// SIMATIC S7-200 project (STEP 7-Micro/WIN), CPU 226 CN REL 02.01

SYMBOL_TABLE ????1
SI1              I0.0     // Sensor de riel
FCI              I0.1     // Final de carrera derecha
FCF              I0.2     // Final de carrera izquierda
SM2B             I0.4     // Sensor de elevamiento vertical
SM2A             I0.3     // Sensor retraido vertical
SAH              I0.5     // Sensor antiHorario de giro
SH               I0.6     // Sensor Horario de giro
SM3B             I0.7     // Sesor extendido horizontal
SM3A             I1.0     // Sensor retraido horizontal
SM4C             I1.1     // Sensor Garra cerrada
                 I1.3     // Alarma servo
SB_2             I2.4     // Pulsador de parada
SB_1             I2.5     // Pulsador de marcha
QS               I2.6     // Zeta de emergencia
SA               I2.7     // Selector de modo
PULSO            Q0.0     // Pulso
DIR              Q0.1     // Direccion
KV2              Q0.3     // Cilndro neumatico vertical
KV1A             Q0.4     // Cilindro rotarorio anti horario
KV1H             Q0.5     // Cilindro rotatorio horario
KV3              Q0.6     // Cilindro doble horizontal
KV4C             Q0.7     // Garra cerrada
KV4A             Q1.0     // Garra abierta
HL1              Q1.5     // Piloto Amarillo
HL2              Q1.6     // Piloto Verde
HL3              Q1.7     // Piloto Rojo
E0               M0.0     // Estado 0
E1               M0.1     // Estado 1
E2               M0.2
E3               M0.3
E4               M0.4
E5               M0.5
E6               M0.6
E7               M0.7
E8               M1.0
E9               M1.1
E10              M1.2
E11              M1.3
E12              M1.4
E13              M1.5
E14              M1.6
E15              M1.7
E16              M2.0
E17              M2.1
E18              M2.2
E19              M2.3
E20              M2.4
E21              M2.5
E22              M2.6
E23              M2.7
EP               M3.0     // Estado de parada momentanea
Marca            M3.1     // Marca auxiliar
EM               M3.2     // Estado de emergencia
SB1_UT           M4.0     // Pulsador de marcha
SB2_UT           M4.1     // Pulsador de parada
QS_UT            M4.2     // Zeta de emergencia
POS_UA           M5.0     // Posicionamiento a la Unidad de Alimentacion
POS_UE           M5.1     // Posicionamiento a la Unidad de Ensamblaje
POS_UP           M5.2     // Posicionamiento a la Unidad de Procesamiento
POS_US           M5.3     // Posicionamiento a la Unidad de Seleccion
END_UA           V0.0     // Finializacion de la Unidad de Alimentacion
END_UE           V12.0    // Finalizacion de la Unidad de Ensamblaje
END_UP           V6.0     // Finalizacion de la Unidad de Procesamiento
END_US           V18.0    // Finalizacion de la Unidad de Seleccion
IN_UA            V3.0     // Iniciar Unidad de Alimentacion
IN_UE            V15.0    // Iniciar Unidad de Ensamblaje
IN_UP            V9.0     // Iniciar Unidad de Procesamiento
IN_US            V21.0    // Iniciar Unidad de Seleccion
                          // UNIDAD DE ALIMENTACION
SB1_UA           M4.3     // Pulsador de marcha
SB2_UA           M4.4     // Pulsador de parada
QS_UA            M4.5     // Zeta de emergencia
KV1_UA           V0.1     // Cilindro neumatico Retenedor
KV2_UA           V0.2     // Cilindro neumatico de empuje
SF_UA            V0.3     // Sensor Fotoelectrico Final
SP_UA            V0.4     // Sensor Fotoelectrico Superior
SP1_UA           V0.5     // Sensor Fotoelectrico Inferior
HL1_UA           V0.6     // Piloto de parada
HL2_UA           V0.7     // Piloto de marcha
HL3_UA           V1.0     // Piloto de emergencia
                          // UNIDAD DE ENSAMBLAJE
SB1_UE           M15.1    // Pulsador de marcha
SB2_UE           M15.2    // Pulsador de parada
QS_UE            M15.3    // Zeta de emergencia
KV1_UE           V12.1    // Cilindro liberador
KV2_UE           V12.2    // Cildro sujetador
KV3_UE           V12.3    // Cilindro rotatorio
KV4_UE           V12.4    // Cilindro vertical
KV5_UE           V12.5    // Cilindro horizontal
KV6_UE           V12.6    // Cilindro de garra
SP1_UE           V13.0    // Sensor del tubo inferior
SP_UE            V13.1    // Sensor del tubo superiro
SST_UE           V13.2    // Sensor salida del tubo
SG_UE            V13.3    // Sensor de recogida de pieza
SF_UE            V13.4    // Sensor de posicion de pieza grande
HL1_UE           V13.5    // Piloto de parada
HL2_UE           V13.6    // Piloto de marcha
HL3_UE           V13.7    // Piloto de emergencia
                          // UNIDAD DE PROCESAMIENTO
SB1_UP           M9.1     // Pulsador de marcha
SB2_UP           M9.2     // Pulsador de parada
QS_UP            M9.3     // Zeta de emergencia
KV1_UP           V6.1     // Cilindro neumatico horizontal
KV2_UP           V6.2     // Cilindro de la pinza
KV3_UP           V6.3     // Cilindro neumatico de compresion
SF1_UP           V6.4     // Sensor optico
HL1_UP           V6.5     // Piloto de parada
HL2_UP           V6.6     // Piloto de marcha
HL3_UP           V6.7     // Piloto de emergencia
                          // UNIDAD DE SELECCION
SB1_US           M21.1    // Pulsador de marcha
SB2_US           M21.2    // Pulsador de parada
QS_US            M21.3    // Zeta de emergencia
KV1_US           V18.1    // Cilindro neumatico 1
KV2_US           V18.2    // Cilindro neumatico 2
KV3_US           V18.3    // Cilindro neumatico 3
motor            V18.4    // Motor
SF_US            V18.5    // Sensor de objetos
SII_US           V18.6    // Sensor inductivo (Metal)
SP_US            V18.7    // Sensor magnetico (plastico)
HL1_US           V19.0    // Piloto de parada
HL2_US           V19.1    // Piloto de marcha
HL3_US           V19.2    // Piloto de emergencia
END_SYMBOL_TABLE

ORGANIZATION_BLOCK PRINCIPAL:OB1
TITLE=????
BEGIN
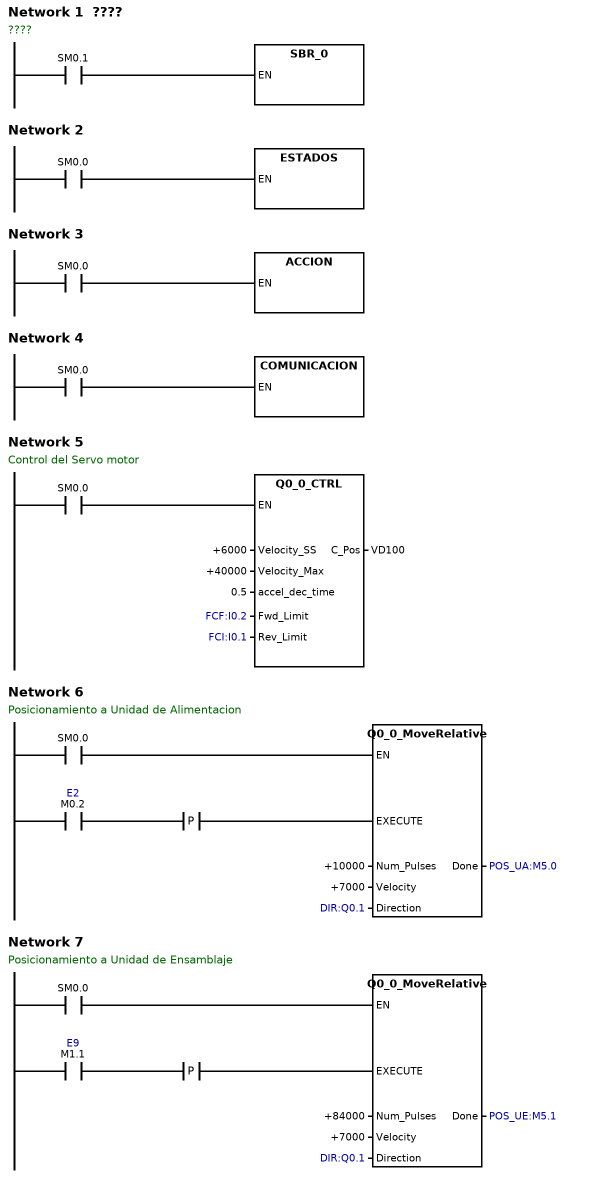
Network 1 // ????
// ????
LD     SM0.1
CALL   SBR_0:SBR0
Network 2
LD     SM0.0
CALL   ESTADOS:SBR1
Network 3
LD     SM0.0
CALL   ACCION:SBR2
Network 4
LD     SM0.0
CALL   COMUNICACION:SBR3
Network 5
// Control del Servo motor
LD     SM0.0
CALL   Q0_0_CTRL:SBR5, +6000, +40000, 0.5, FCF:I0.2, FCI:I0.1, VD100
Network 6
// Posicionamiento a Unidad de Alimentacion
LD     SM0.0
=      L60.0
LD     E2:M0.2
EU
=      L63.7
LD     L60.0
CALL   Q0_0_MoveRelative:SBR8, L63.7, +10000, +7000, DIR:Q0.1, POS_UA:M5.0
Network 7
// Posicionamiento a Unidad de Ensamblaje
LD     SM0.0
=      L60.0
LD     E9:M1.1
EU
=      L63.7
LD     L60.0
CALL   Q0_0_MoveRelative:SBR8, L63.7, +84000, +7000, DIR:Q0.1, POS_UE:M5.1
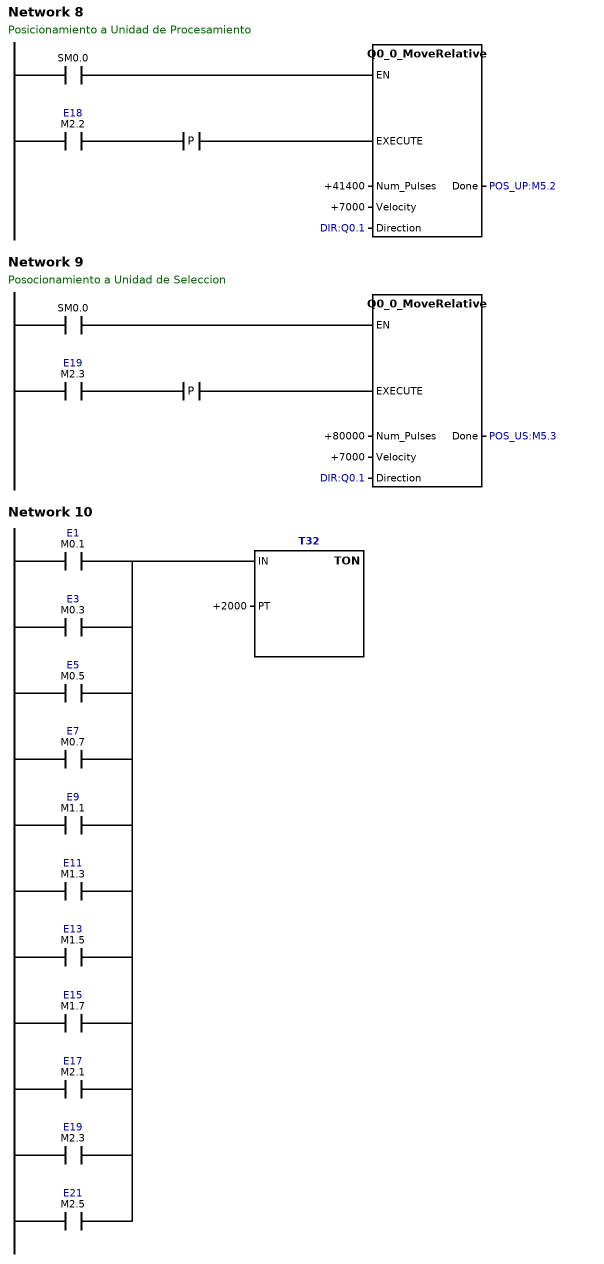
Network 8
// Posicionamiento a Unidad de Procesamiento
LD     SM0.0
=      L60.0
LD     E18:M2.2
EU
=      L63.7
LD     L60.0
CALL   Q0_0_MoveRelative:SBR8, L63.7, +41400, +7000, DIR:Q0.1, POS_UP:M5.2
Network 9
// Posocionamiento a Unidad de Seleccion
LD     SM0.0
=      L60.0
LD     E19:M2.3
EU
=      L63.7
LD     L60.0
CALL   Q0_0_MoveRelative:SBR8, L63.7, +80000, +7000, DIR:Q0.1, POS_US:M5.3
Network 10
LD     E1:M0.1
O      E3:M0.3
O      E5:M0.5
O      E7:M0.7
O      E9:M1.1
O      E11:M1.3
O      E13:M1.5
O      E15:M1.7
O      E17:M2.1
O      E19:M2.3
O      E21:M2.5
TON    T32, +2000
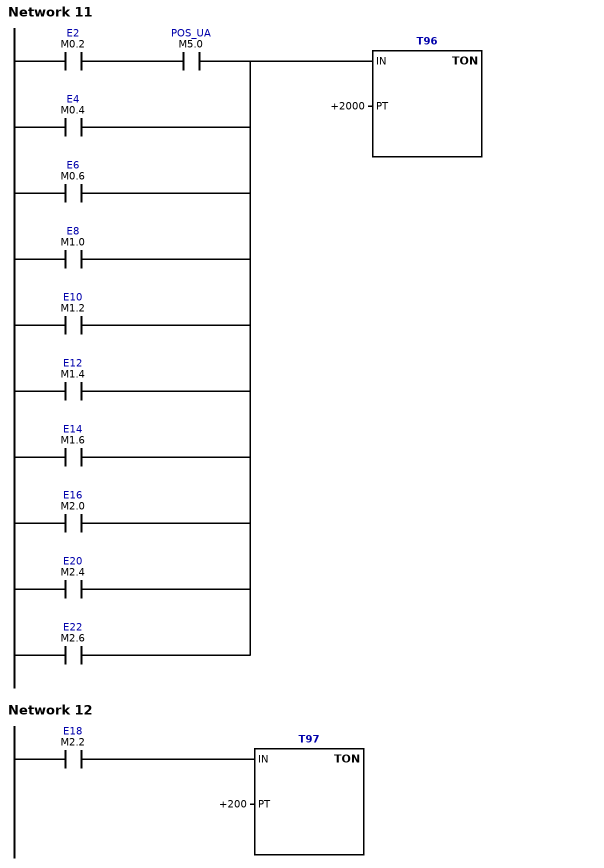
Network 11
LD     E2:M0.2
A      POS_UA:M5.0
O      E4:M0.4
O      E6:M0.6
O      E8:M1.0
O      E10:M1.2
O      E12:M1.4
O      E14:M1.6
O      E16:M2.0
O      E20:M2.4
O      E22:M2.6
TON    T96, +2000
Network 12
LD     E18:M2.2
TON    T97, +200
END_ORGANIZATION_BLOCK

SUBROUTINE_BLOCK SBR_0:SBR0
TITLE=?????
BEGIN
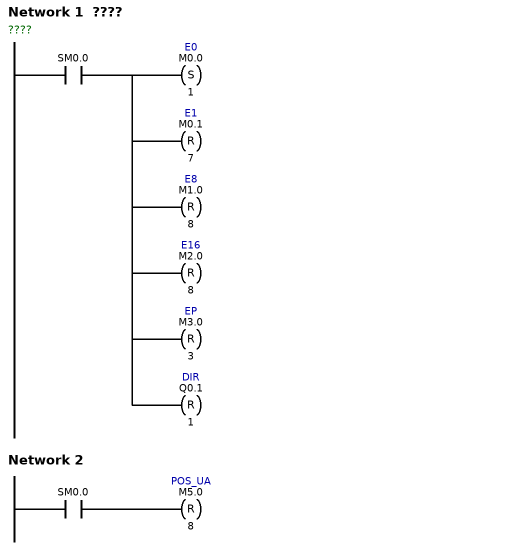
Network 1 // ????
// ????
LD     SM0.0
S      E0:M0.0, 1
R      E1:M0.1, 7
R      E8:M1.0, 8
R      E16:M2.0, 8
R      EP:M3.0, 3
R      DIR:Q0.1, 1
Network 2
LD     SM0.0
R      POS_UA:M5.0, 8
END_SUBROUTINE_BLOCK

SUBROUTINE_BLOCK ESTADOS:SBR1
TITLE=
BEGIN
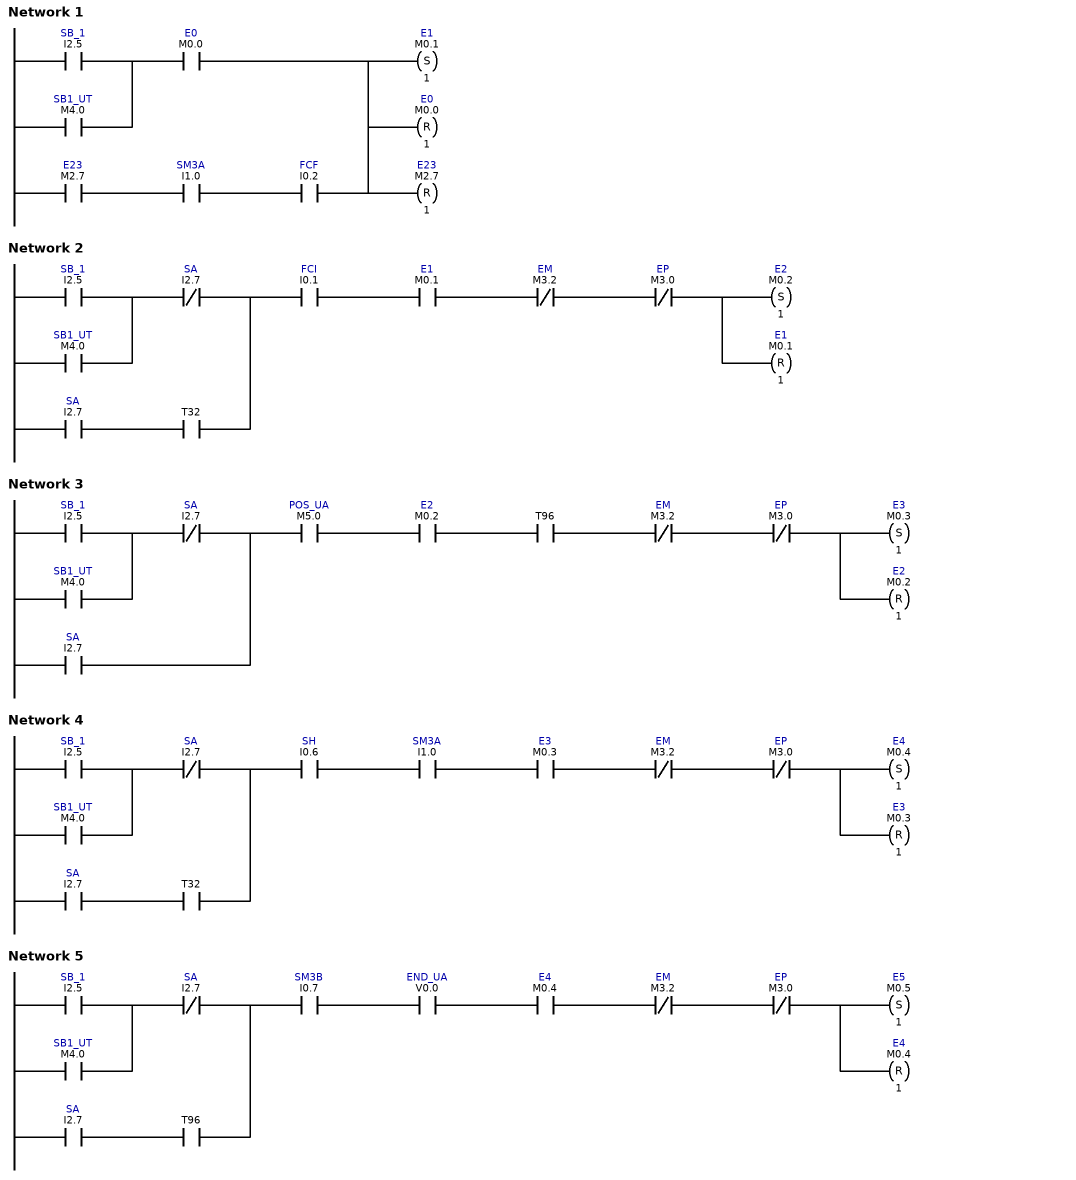
Network 1
LD     SB_1:I2.5
O      SB1_UT:M4.0
A      E0:M0.0
LD     E23:M2.7
A      SM3A:I1.0
A      FCF:I0.2
OLD
S      E1:M0.1, 1
R      E0:M0.0, 1
R      E23:M2.7, 1
Network 2
LD     SB_1:I2.5
O      SB1_UT:M4.0
AN     SA:I2.7
LD     SA:I2.7
A      T32
OLD
A      FCI:I0.1
A      E1:M0.1
AN     EM:M3.2
AN     EP:M3.0
S      E2:M0.2, 1
R      E1:M0.1, 1
Network 3
LD     SB_1:I2.5
O      SB1_UT:M4.0
AN     SA:I2.7
O      SA:I2.7
A      POS_UA:M5.0
A      E2:M0.2
A      T96
AN     EM:M3.2
AN     EP:M3.0
S      E3:M0.3, 1
R      E2:M0.2, 1
Network 4
LD     SB_1:I2.5
O      SB1_UT:M4.0
AN     SA:I2.7
LD     SA:I2.7
A      T32
OLD
A      SH:I0.6
A      SM3A:I1.0
A      E3:M0.3
AN     EM:M3.2
AN     EP:M3.0
S      E4:M0.4, 1
R      E3:M0.3, 1
Network 5
LD     SB_1:I2.5
O      SB1_UT:M4.0
AN     SA:I2.7
LD     SA:I2.7
A      T96
OLD
A      SM3B:I0.7
A      END_UA:V0.0
A      E4:M0.4
AN     EM:M3.2
AN     EP:M3.0
S      E5:M0.5, 1
R      E4:M0.4, 1
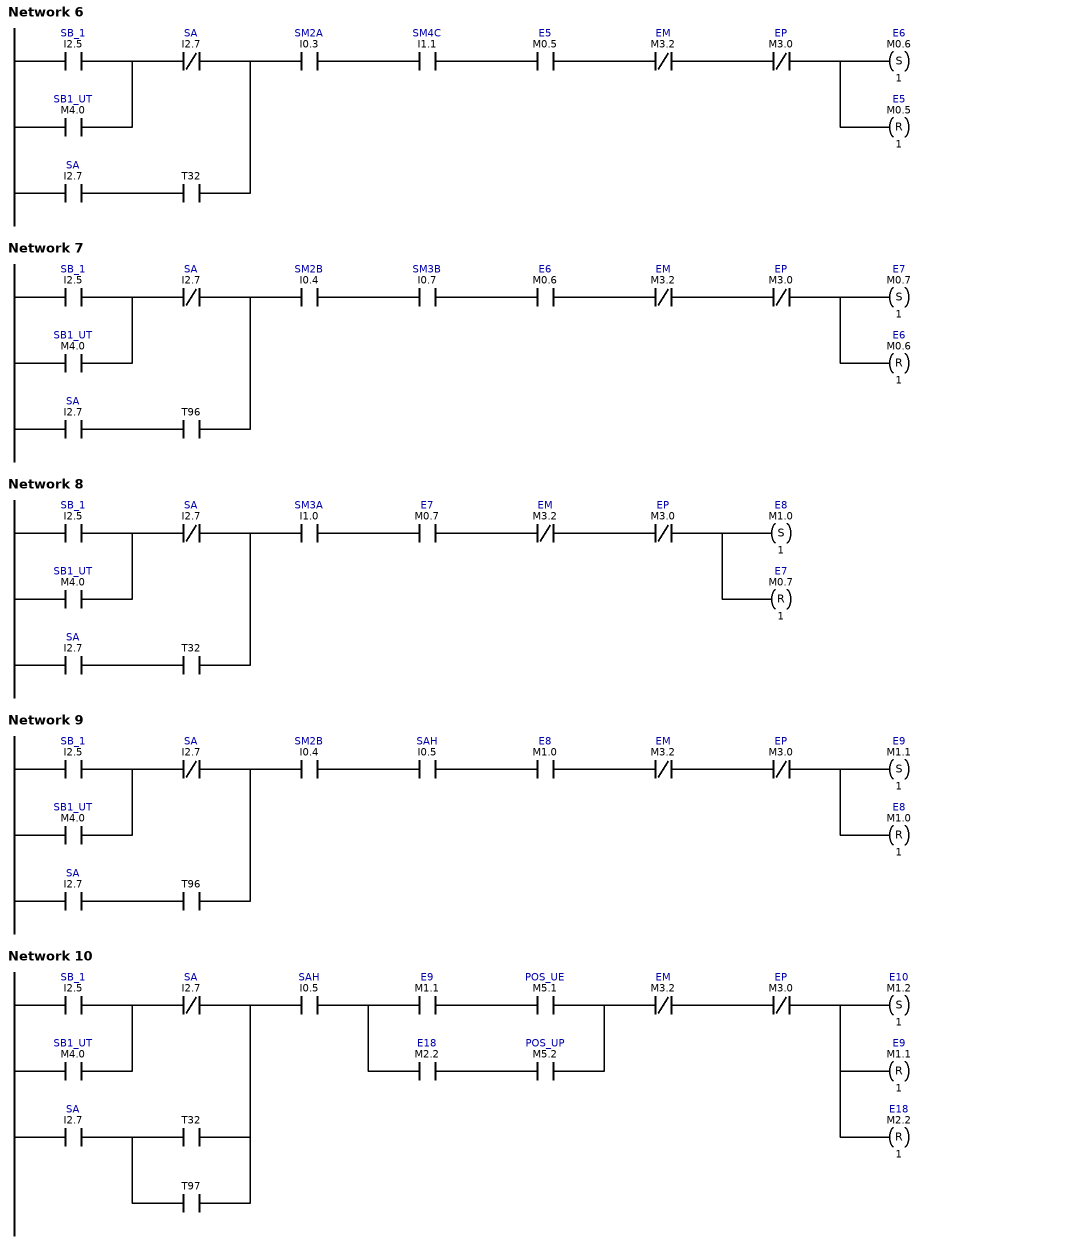
Network 6
LD     SB_1:I2.5
O      SB1_UT:M4.0
AN     SA:I2.7
LD     SA:I2.7
A      T32
OLD
A      SM2A:I0.3
A      SM4C:I1.1
A      E5:M0.5
AN     EM:M3.2
AN     EP:M3.0
S      E6:M0.6, 1
R      E5:M0.5, 1
Network 7
LD     SB_1:I2.5
O      SB1_UT:M4.0
AN     SA:I2.7
LD     SA:I2.7
A      T96
OLD
A      SM2B:I0.4
A      SM3B:I0.7
A      E6:M0.6
AN     EM:M3.2
AN     EP:M3.0
S      E7:M0.7, 1
R      E6:M0.6, 1
Network 8
LD     SB_1:I2.5
O      SB1_UT:M4.0
AN     SA:I2.7
LD     SA:I2.7
A      T32
OLD
A      SM3A:I1.0
A      E7:M0.7
AN     EM:M3.2
AN     EP:M3.0
S      E8:M1.0, 1
R      E7:M0.7, 1
Network 9
LD     SB_1:I2.5
O      SB1_UT:M4.0
AN     SA:I2.7
LD     SA:I2.7
A      T96
OLD
A      SM2B:I0.4
A      SAH:I0.5
A      E8:M1.0
AN     EM:M3.2
AN     EP:M3.0
S      E9:M1.1, 1
R      E8:M1.0, 1
Network 10
LD     SB_1:I2.5
O      SB1_UT:M4.0
AN     SA:I2.7
LD     SA:I2.7
LD     T32
O      T97
ALD
OLD
A      SAH:I0.5
LD     E9:M1.1
A      POS_UE:M5.1
LD     E18:M2.2
A      POS_UP:M5.2
OLD
ALD
AN     EM:M3.2
AN     EP:M3.0
S      E10:M1.2, 1
R      E9:M1.1, 1
R      E18:M2.2, 1
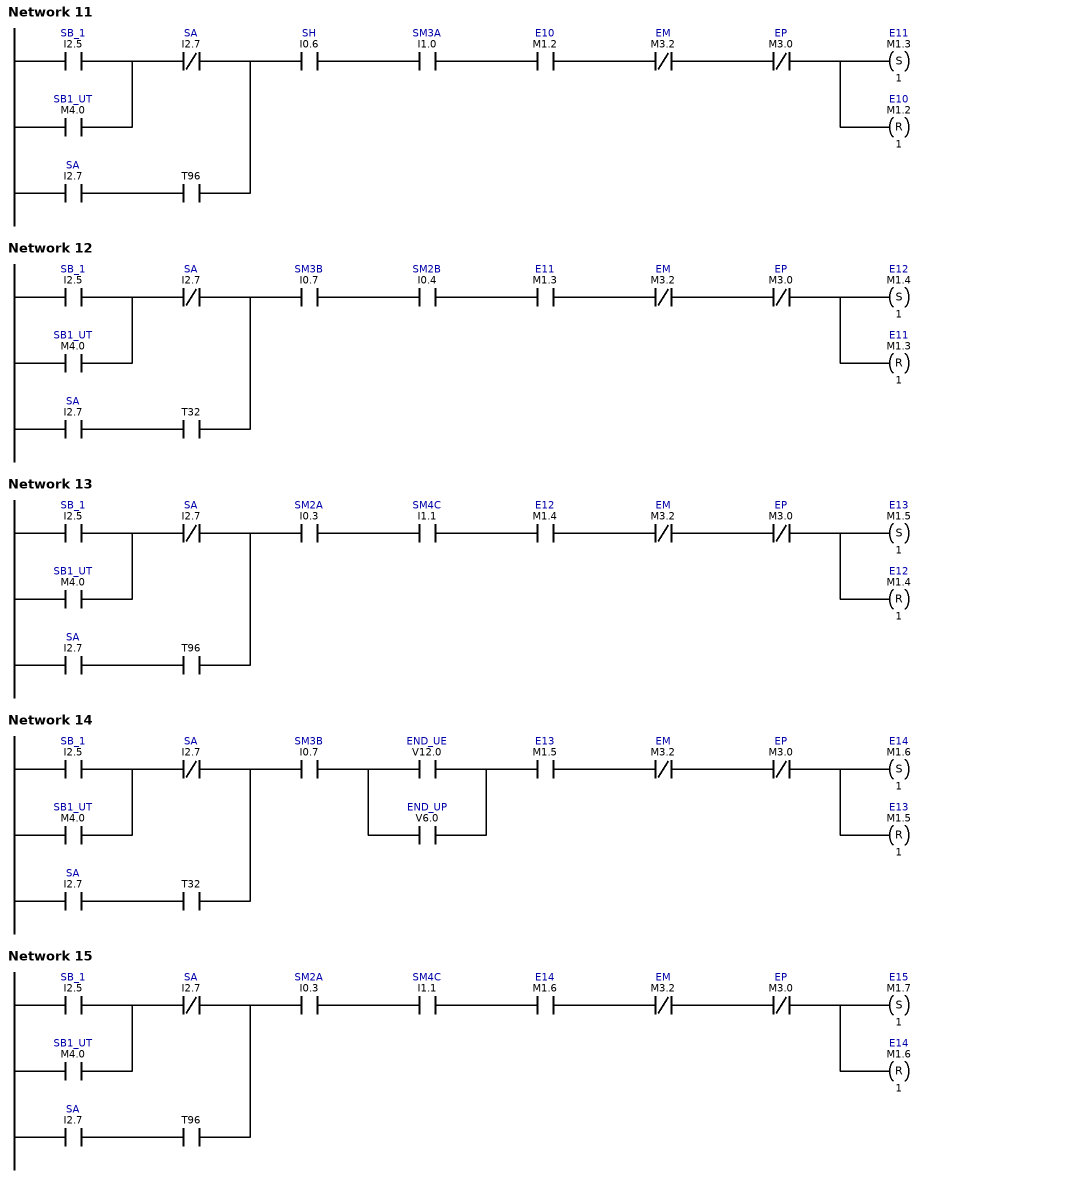
Network 11
LD     SB_1:I2.5
O      SB1_UT:M4.0
AN     SA:I2.7
LD     SA:I2.7
A      T96
OLD
A      SH:I0.6
A      SM3A:I1.0
A      E10:M1.2
AN     EM:M3.2
AN     EP:M3.0
S      E11:M1.3, 1
R      E10:M1.2, 1
Network 12
LD     SB_1:I2.5
O      SB1_UT:M4.0
AN     SA:I2.7
LD     SA:I2.7
A      T32
OLD
A      SM3B:I0.7
A      SM2B:I0.4
A      E11:M1.3
AN     EM:M3.2
AN     EP:M3.0
S      E12:M1.4, 1
R      E11:M1.3, 1
Network 13
LD     SB_1:I2.5
O      SB1_UT:M4.0
AN     SA:I2.7
LD     SA:I2.7
A      T96
OLD
A      SM2A:I0.3
A      SM4C:I1.1
A      E12:M1.4
AN     EM:M3.2
AN     EP:M3.0
S      E13:M1.5, 1
R      E12:M1.4, 1
Network 14
LD     SB_1:I2.5
O      SB1_UT:M4.0
AN     SA:I2.7
LD     SA:I2.7
A      T32
OLD
A      SM3B:I0.7
LD     END_UE:V12.0
O      END_UP:V6.0
ALD
A      E13:M1.5
AN     EM:M3.2
AN     EP:M3.0
S      E14:M1.6, 1
R      E13:M1.5, 1
Network 15
LD     SB_1:I2.5
O      SB1_UT:M4.0
AN     SA:I2.7
LD     SA:I2.7
A      T96
OLD
A      SM2A:I0.3
A      SM4C:I1.1
A      E14:M1.6
AN     EM:M3.2
AN     EP:M3.0
S      E15:M1.7, 1
R      E14:M1.6, 1
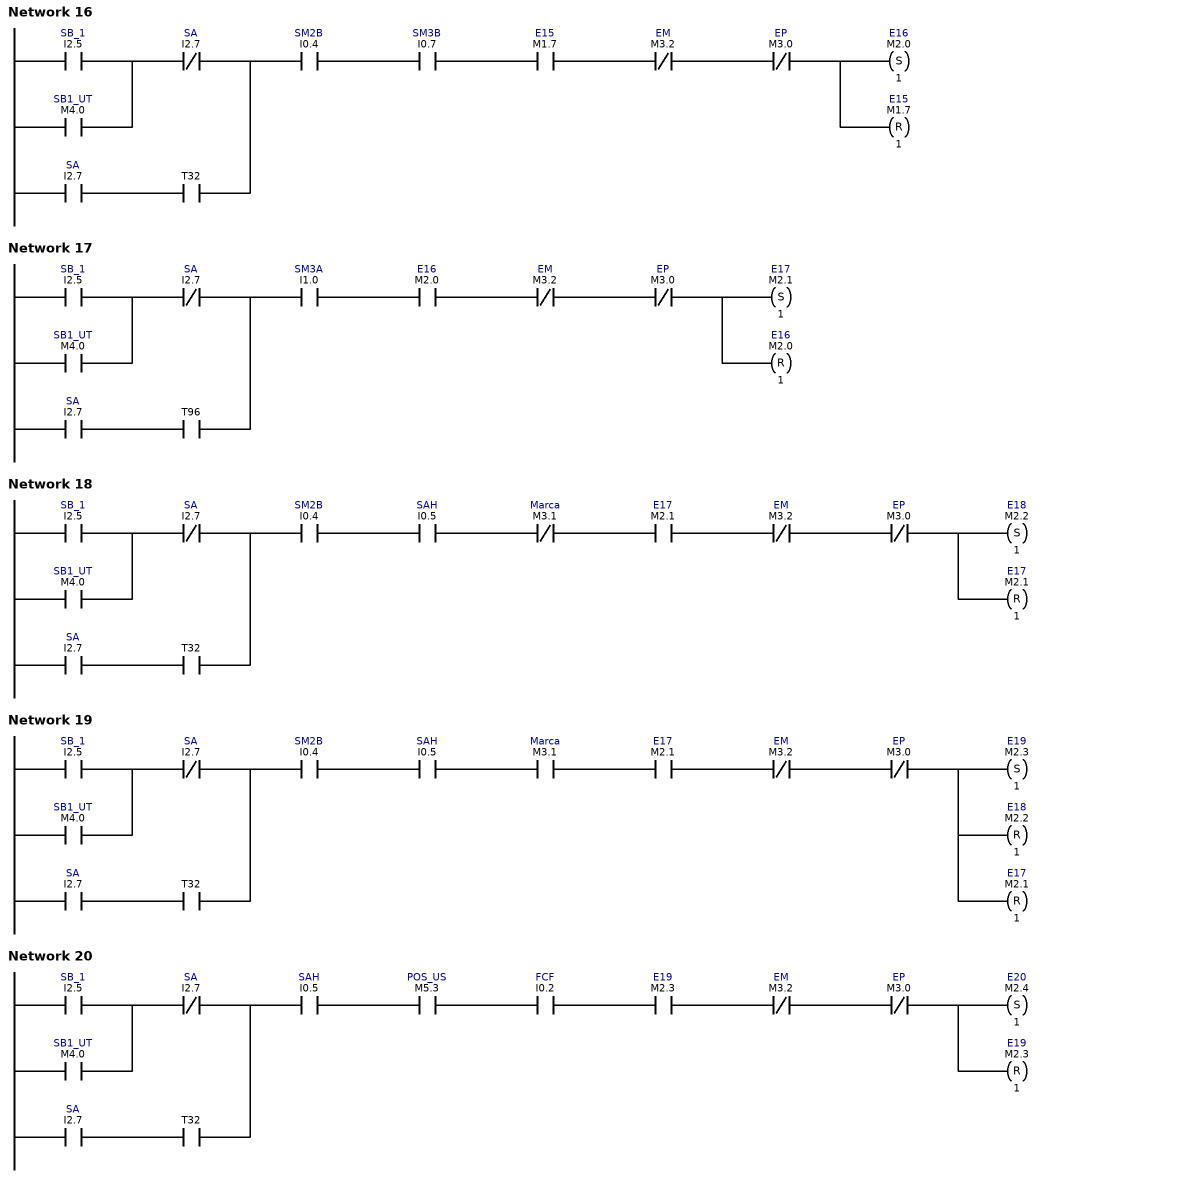
Network 16
LD     SB_1:I2.5
O      SB1_UT:M4.0
AN     SA:I2.7
LD     SA:I2.7
A      T32
OLD
A      SM2B:I0.4
A      SM3B:I0.7
A      E15:M1.7
AN     EM:M3.2
AN     EP:M3.0
S      E16:M2.0, 1
R      E15:M1.7, 1
Network 17
LD     SB_1:I2.5
O      SB1_UT:M4.0
AN     SA:I2.7
LD     SA:I2.7
A      T96
OLD
A      SM3A:I1.0
A      E16:M2.0
AN     EM:M3.2
AN     EP:M3.0
S      E17:M2.1, 1
R      E16:M2.0, 1
Network 18
LD     SB_1:I2.5
O      SB1_UT:M4.0
AN     SA:I2.7
LD     SA:I2.7
A      T32
OLD
A      SM2B:I0.4
A      SAH:I0.5
AN     Marca:M3.1
A      E17:M2.1
AN     EM:M3.2
AN     EP:M3.0
S      E18:M2.2, 1
R      E17:M2.1, 1
Network 19
LD     SB_1:I2.5
O      SB1_UT:M4.0
AN     SA:I2.7
LD     SA:I2.7
A      T32
OLD
A      SM2B:I0.4
A      SAH:I0.5
A      Marca:M3.1
A      E17:M2.1
AN     EM:M3.2
AN     EP:M3.0
S      E19:M2.3, 1
R      E18:M2.2, 1
R      E17:M2.1, 1
Network 20
LD     SB_1:I2.5
O      SB1_UT:M4.0
AN     SA:I2.7
LD     SA:I2.7
A      T32
OLD
A      SAH:I0.5
A      POS_US:M5.3
A      FCF:I0.2
A      E19:M2.3
AN     EM:M3.2
AN     EP:M3.0
S      E20:M2.4, 1
R      E19:M2.3, 1
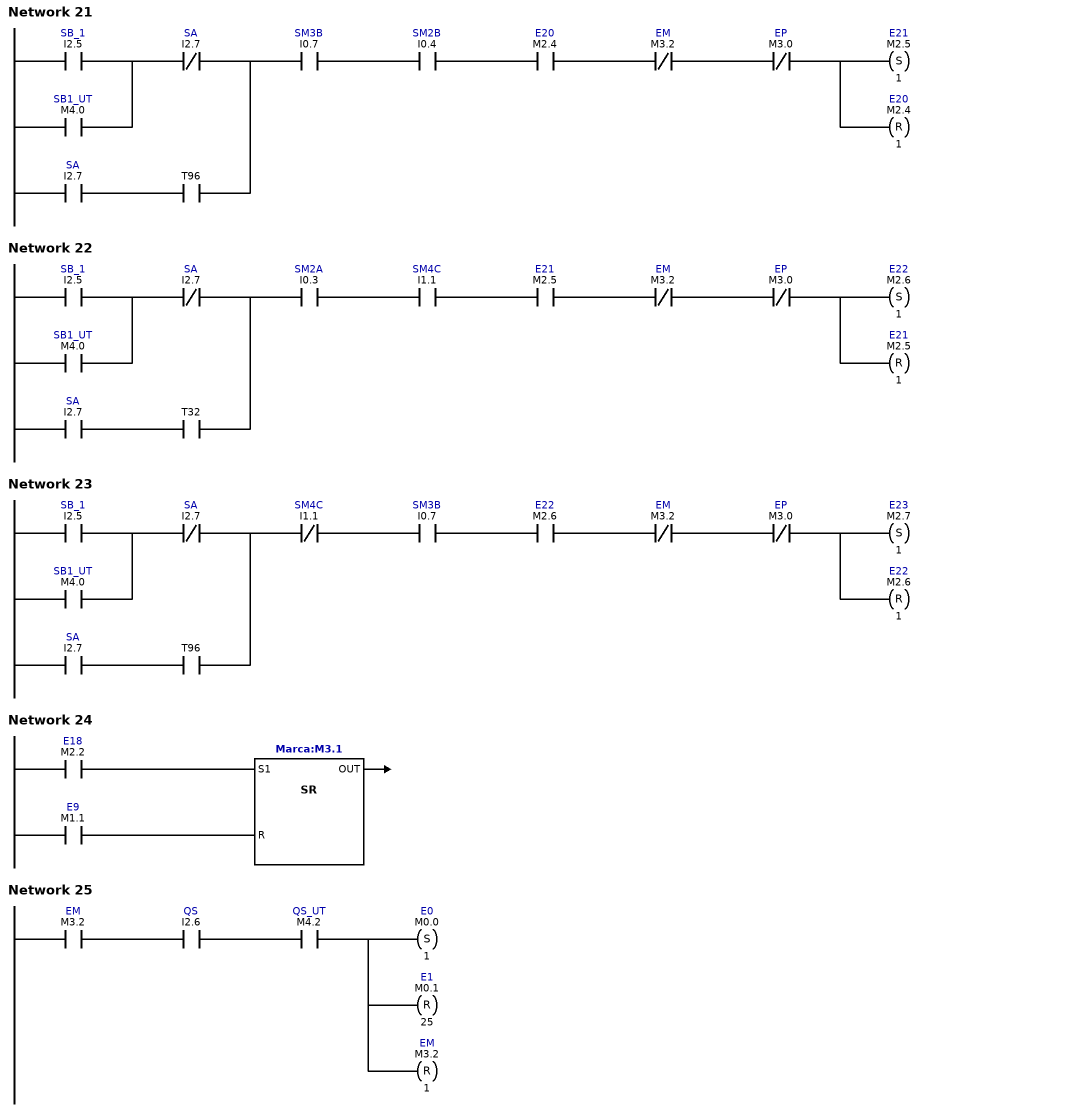
Network 21
LD     SB_1:I2.5
O      SB1_UT:M4.0
AN     SA:I2.7
LD     SA:I2.7
A      T96
OLD
A      SM3B:I0.7
A      SM2B:I0.4
A      E20:M2.4
AN     EM:M3.2
AN     EP:M3.0
S      E21:M2.5, 1
R      E20:M2.4, 1
Network 22
LD     SB_1:I2.5
O      SB1_UT:M4.0
AN     SA:I2.7
LD     SA:I2.7
A      T32
OLD
A      SM2A:I0.3
A      SM4C:I1.1
A      E21:M2.5
AN     EM:M3.2
AN     EP:M3.0
S      E22:M2.6, 1
R      E21:M2.5, 1
Network 23
LD     SB_1:I2.5
O      SB1_UT:M4.0
AN     SA:I2.7
LD     SA:I2.7
A      T96
OLD
AN     SM4C:I1.1
A      SM3B:I0.7
A      E22:M2.6
AN     EM:M3.2
AN     EP:M3.0
S      E23:M2.7, 1
R      E22:M2.6, 1
Network 24
LD     E18:M2.2
LD     E9:M1.1
NOT
A      Marca:M3.1
OLD
=      Marca:M3.1
Network 25
LD     EM:M3.2
A      QS:I2.6
A      QS_UT:M4.2
S      E0:M0.0, 1
R      E1:M0.1, 25
R      EM:M3.2, 1
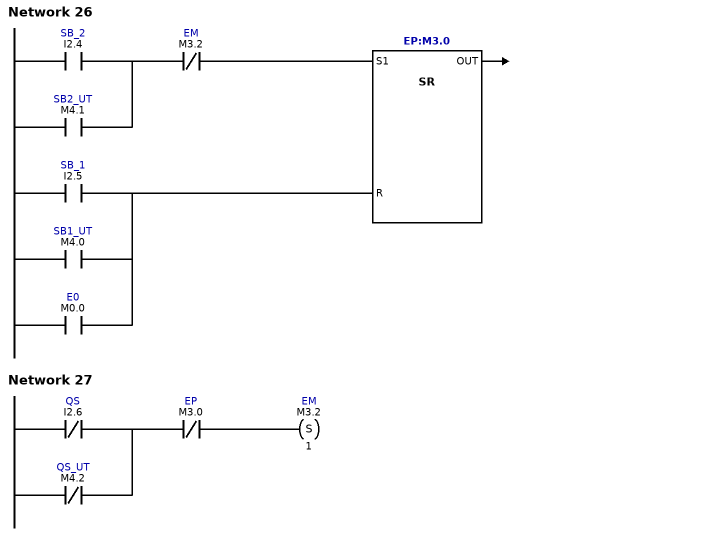
Network 26
LD     SB_2:I2.4
O      SB2_UT:M4.1
AN     EM:M3.2
LD     SB_1:I2.5
O      SB1_UT:M4.0
O      E0:M0.0
NOT
A      EP:M3.0
OLD
=      EP:M3.0
Network 27
LDN    QS:I2.6
ON     QS_UT:M4.2
AN     EP:M3.0
S      EM:M3.2, 1
END_SUBROUTINE_BLOCK

SUBROUTINE_BLOCK ACCION:SBR2
TITLE=
BEGIN
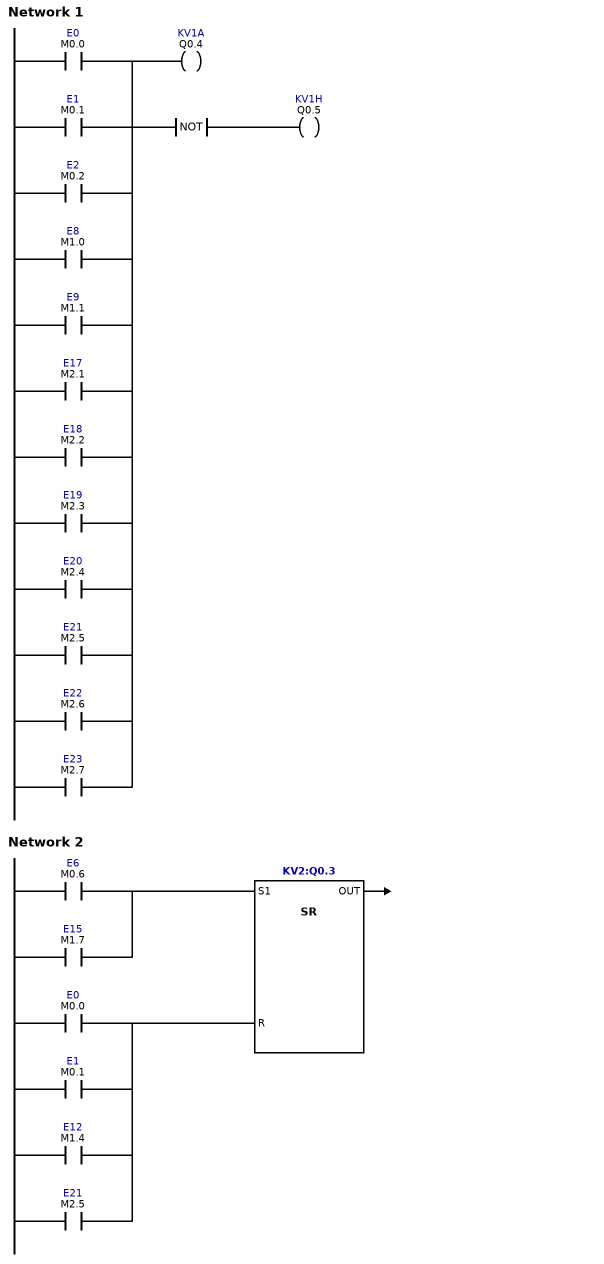
Network 1
LD     E0:M0.0
O      E1:M0.1
O      E2:M0.2
O      E8:M1.0
O      E9:M1.1
O      E17:M2.1
O      E18:M2.2
O      E19:M2.3
O      E20:M2.4
O      E21:M2.5
O      E22:M2.6
O      E23:M2.7
=      KV1A:Q0.4
NOT
=      KV1H:Q0.5
Network 2
LD     E6:M0.6
O      E15:M1.7
LD     E0:M0.0
O      E1:M0.1
O      E12:M1.4
O      E21:M2.5
NOT
A      KV2:Q0.3
OLD
=      KV2:Q0.3
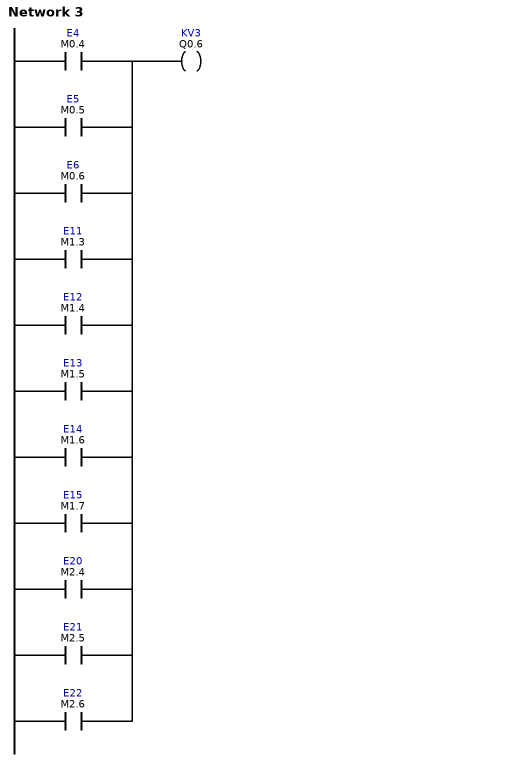
Network 3
LD     E4:M0.4
O      E5:M0.5
O      E6:M0.6
O      E11:M1.3
O      E12:M1.4
O      E13:M1.5
O      E14:M1.6
O      E15:M1.7
O      E20:M2.4
O      E21:M2.5
O      E22:M2.6
=      KV3:Q0.6
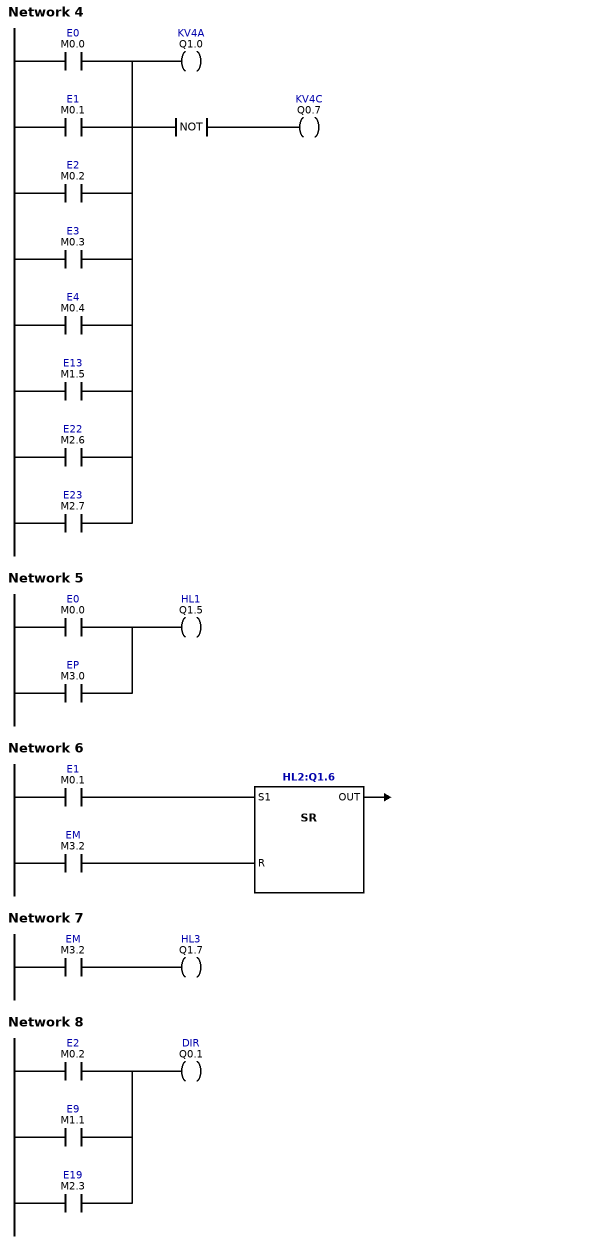
Network 4
LD     E0:M0.0
O      E1:M0.1
O      E2:M0.2
O      E3:M0.3
O      E4:M0.4
O      E13:M1.5
O      E22:M2.6
O      E23:M2.7
=      KV4A:Q1.0
NOT
=      KV4C:Q0.7
Network 5
LD     E0:M0.0
O      EP:M3.0
=      HL1:Q1.5
Network 6
LD     E1:M0.1
LD     EM:M3.2
NOT
A      HL2:Q1.6
OLD
=      HL2:Q1.6
Network 7
LD     EM:M3.2
=      HL3:Q1.7
Network 8
LD     E2:M0.2
O      E9:M1.1
O      E19:M2.3
=      DIR:Q0.1
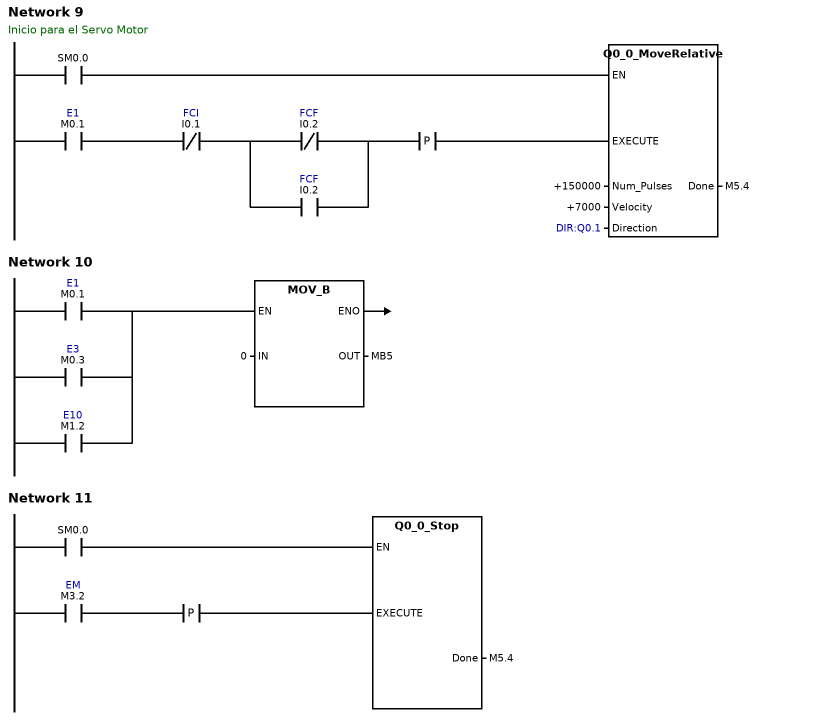
Network 9
// Inicio para el Servo Motor
LD     SM0.0
=      L60.0
LD     E1:M0.1
AN     FCI:I0.1
LDN    FCF:I0.2
O      FCF:I0.2
ALD
EU
=      L63.7
LD     L60.0
CALL   Q0_0_MoveRelative:SBR8, L63.7, +150000, +7000, DIR:Q0.1, M5.4
Network 10
LD     E1:M0.1
O      E3:M0.3
O      E10:M1.2
MOVB   0, MB5
Network 11
LD     SM0.0
=      L60.0
LD     EM:M3.2
EU
=      L63.7
LD     L60.0
CALL   Q0_0_Stop:SBR10, L63.7, M5.4
END_SUBROUTINE_BLOCK

SUBROUTINE_BLOCK COMUNICACION:SBR3
TITLE=
BEGIN
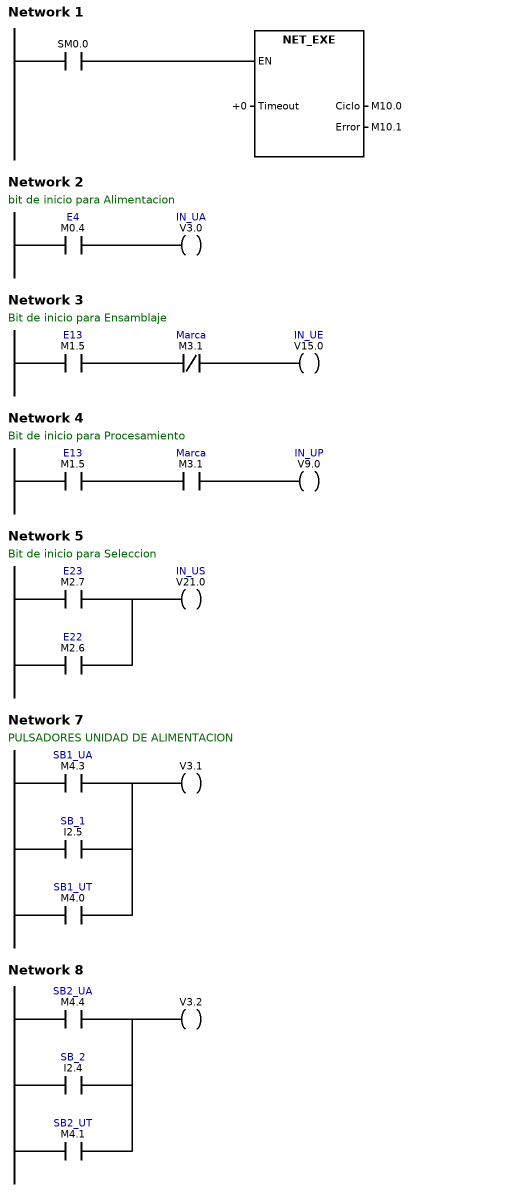
Network 1
LD     SM0.0
CALL   NET_EXE:SBR4, +0, M10.0, M10.1
Network 2
// bit de inicio para Alimentacion 
LD     E4:M0.4
=      IN_UA:V3.0
Network 3
// Bit de inicio para Ensamblaje
LD     E13:M1.5
AN     Marca:M3.1
=      IN_UE:V15.0
Network 4
// Bit de inicio para Procesamiento
LD     E13:M1.5
A      Marca:M3.1
=      IN_UP:V9.0
Network 5
// Bit de inicio para Seleccion
LD     E23:M2.7
O      E22:M2.6
=      IN_US:V21.0
Network 6
// PULSADORES
Network 7
// PULSADORES UNIDAD DE ALIMENTACION
LD     SB1_UA:M4.3
O      SB_1:I2.5
O      SB1_UT:M4.0
=      V3.1
Network 8
LD     SB2_UA:M4.4
O      SB_2:I2.4
O      SB2_UT:M4.1
=      V3.2
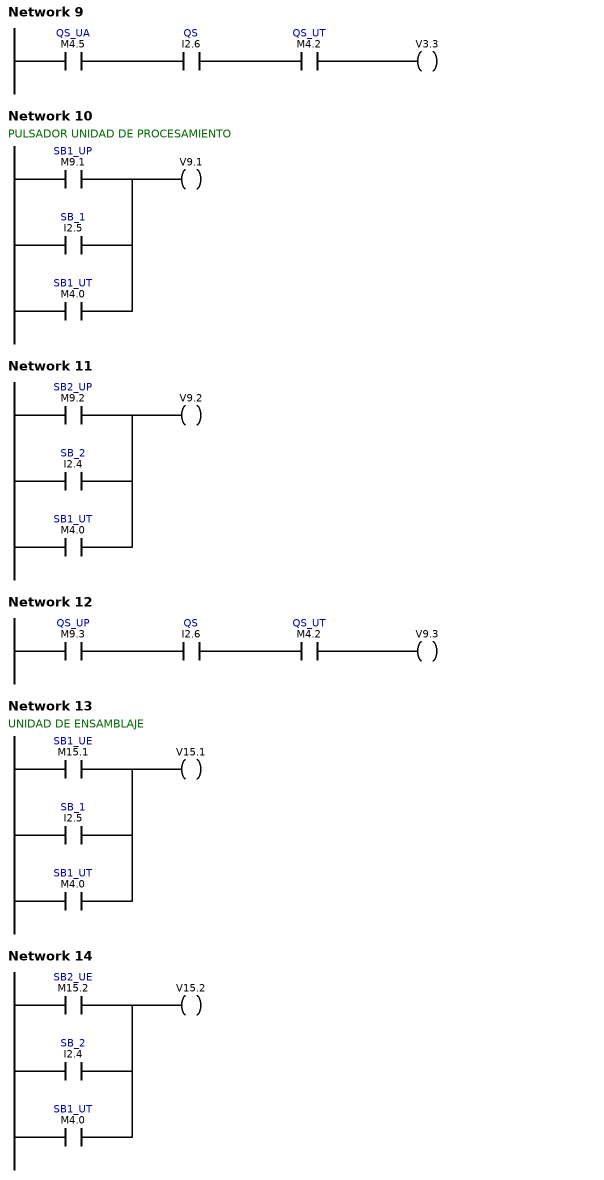
Network 9
LD     QS_UA:M4.5
A      QS:I2.6
A      QS_UT:M4.2
=      V3.3
Network 10
// PULSADOR UNIDAD DE PROCESAMIENTO
LD     SB1_UP:M9.1
O      SB_1:I2.5
O      SB1_UT:M4.0
=      V9.1
Network 11
LD     SB2_UP:M9.2
O      SB_2:I2.4
O      SB1_UT:M4.0
=      V9.2
Network 12
LD     QS_UP:M9.3
A      QS:I2.6
A      QS_UT:M4.2
=      V9.3
Network 13
// UNIDAD DE ENSAMBLAJE
LD     SB1_UE:M15.1
O      SB_1:I2.5
O      SB1_UT:M4.0
=      V15.1
Network 14
LD     SB2_UE:M15.2
O      SB_2:I2.4
O      SB1_UT:M4.0
=      V15.2
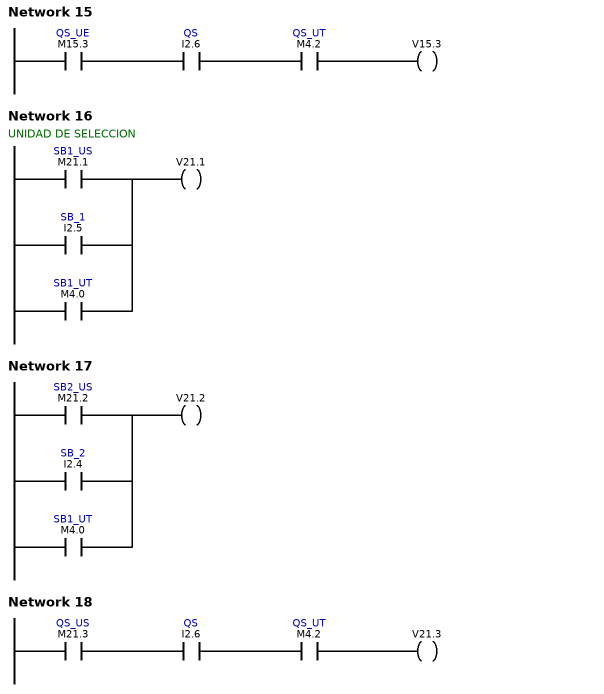
Network 15
LD     QS_UE:M15.3
A      QS:I2.6
A      QS_UT:M4.2
=      V15.3
Network 16
// UNIDAD DE SELECCION
LD     SB1_US:M21.1
O      SB_1:I2.5
O      SB1_UT:M4.0
=      V21.1
Network 17
LD     SB2_US:M21.2
O      SB_2:I2.4
O      SB1_UT:M4.0
=      V21.2
Network 18
LD     QS_US:M21.3
A      QS:I2.6
A      QS_UT:M4.2
=      V21.3
END_SUBROUTINE_BLOCK

// SBR4: protected block, not included

// SBR5: protected block, not included

// SBR6: protected block, not included

// SBR7: protected block, not included

// SBR8: protected block, not included

// SBR9: protected block, not included

// SBR10: protected block, not included

// INT1: protected block, not included

// INT2: protected block, not included

// INT3: protected block, not included
